Fanuc KAREL source: ko00056.KL

-- PROVISIONAL review KL for V770-1; original PC SHA256 34b3d25996f86458edb842b66256344e34ebbd06ee8caa1f7d185ea333aca624
-- Incomplete behavior may be omitted. Consult companion uncertainty JSON. Do not deploy.
PROGRAM KO00056
%NOLOCKGROUP
BEGIN
  -- UNRESOLVED_PC offsets 5-12; opcodes 9D,23
  -- UNRESOLVED_PC offsets 17-69; opcodes 27,27,49,7E,AD,27,49,7E,AD,22,31,7E,4A
  -- UNRESOLVED_PC offsets 74-78; opcodes 7F
END KO00056
